(* IEC 61131-3 sources: axsharp/src/AXSharp.connectors/tests/ax-test-project/src, 12 files *)

(* ---- enum.st ---- *)
TYPE
    Colors : (RED, GREEN, BLUE);
END_TYPE

(* ---- complexArrayItem.st ---- *)
{S7.extern=ReadWrite}
CLASS complexArrayItem
    VAR PUBLIC
        itemBOOL	        :       BOOL	      ;
        itemSTRING	        :   STRING	      ;
        itemINT	    :       INT	      ;

    END_VAR
END_CLASS

(* ---- complexArrayItemNested.st ---- *)
{S7.extern=ReadWrite}
CLASS complexArrayItemNested
    VAR PUBLIC
        nesteditemBOOL	        :       BOOL	      ;
        nesteditemSTRING	        :   STRING	      ;
        nesteditemINT	    :       INT	      ;
        nestedComplex: complexArrayItem;
    END_VAR
END_CLASS

(* ---- full_of_primitives.st ---- *)
{S7.extern=ReadWrite}
CLASS full_of_primitives
    VAR PUBLIC
        myBOOL	        :       BOOL	      ;
        myBYTE	        :       BYTE	      ;
        myWORD	        :       WORD	      ;
        myDWORD	        :       DWORD	      ;
        myLWORD	        :       LWORD	      ;
        mySINT	        :       SINT	      ;
        myINT	          :       INT	        ;
        myDINT	        :       DINT	      ;
        myLINT	        :       LINT	      ;
        myUSINT	        :       USINT	      ;
        myUINT	        :       UINT	      ;
        myUDINT	        :       UDINT	      ;
        myULINT	        :       ULINT	      ;
        myREAL	        :       REAL	      ;
        myLREAL	        :       LREAL	      ;
        myTIME	        :       TIME	      ;
        myLTIME	        :       LTIME	      ;
        myDATE	        :       DATE	      ;
        myLDATE	        :       LDATE	      ;
        myTIME_OF_DAY	:       TIME_OF_DAY	  ;
        myLTIME_OF_DAY	:       LTIME_OF_DAY  ;
        myDATE_AND_TIME  :      DATE_AND_TIME ;
        myLDATE_AND_TIME :      LDATE_AND_TIME;
        myCHAR	        :       CHAR	      ;
        myWCHAR	        :       WCHAR	      ;
         mySTRING	        :   STRING	      ;
         myWSTRING	    :       WSTRING	      ;
    END_VAR
END_CLASS

(* ---- full_of_primitives_match.st ---- *)
{S7.extern=ReadWrite}
CLASS full_of_primitives_match
    VAR PUBLIC

        myBOOL	            : BOOL;
        myBYTE	            : BOOL;
        myWORD	            : BOOL;
        myDWORD	        : BOOL;
        myLWORD	        : BOOL;
        mySINT	            : BOOL;
        myINT	            : BOOL;
        myDINT	            : BOOL;
        myLINT	            : BOOL;
        myUSINT	        : BOOL;
        myUINT	            : BOOL;
        myUDINT	        : BOOL;
        myULINT	        : BOOL;
        myREAL	            : BOOL;
        myLREAL	        : BOOL;
        myTIME	            : BOOL;
        myLTIME	        : BOOL;
        myDATE	            : BOOL;
        myLDATE	        : BOOL;
        myTIME_OF_DAY	    : BOOL;
        myLTIME_OF_DAY	    : BOOL;
        myDATE_AND_TIME    : BOOL;
        myLDATE_AND_TIME   : BOOL;
        myCHAR	            : BOOL;
        myWCHAR	        : BOOL;
        mySTRING	        : BOOL;
        myWSTRING	        : BOOL;
    END_VAR
END_CLASS

(* ---- hierarchy.st ---- *)
{S7.extern=ReadWrite}
CLASS hierarchy
    VAR PUBLIC
        item  :      hierarchy_2;
    END_VAR
END_CLASS

(* ---- hierarchy_0.st ---- *)
{S7.extern=ReadWrite}
CLASS hierarchy_0
    VAR PUBLIC
        item_member_property_1   :     full_of_primitives;
        item_member_property_2   :     full_of_primitives;
        item_member_property_3   :     full_of_primitives;
        item_member_property_4   :     full_of_primitives;
        item_member_property_5   :     full_of_primitives;
        item_member_property_6   :     full_of_primitives;
        item_member_property_7   :     full_of_primitives;
        item_member_property_8   :     full_of_primitives;
        item_member_property_9   :     full_of_primitives;
        item_member_property_10  :     full_of_primitives;
        item_member_property_12  :     full_of_primitives;
        item_member_property_13  :     full_of_primitives;
        item_member_property_14  :     full_of_primitives;
        item_member_property_15  :     full_of_primitives;
        item_member_property_16  :     full_of_primitives;
        item_member_property_17  :     full_of_primitives;
        item_member_property_18  :     full_of_primitives;
        item_member_property_19  :     full_of_primitives;
    END_VAR
END_CLASS

(* ---- hierarchy_2.st ---- *)
{S7.extern=ReadWrite}
CLASS hierarchy_2
    VAR PUBLIC
        item_member_property_1   :     hierarchy_0;
        item_member_property_2   :     hierarchy_0;
        item_member_property_3   :     hierarchy_0;
        item_member_property_4   :     hierarchy_0;
        item_member_property_5   :     hierarchy_0;
        item_member_property_6   :     hierarchy_0;
        item_member_property_7   :     hierarchy_0;
        item_member_property_8   :     hierarchy_0;
        item_member_property_9   :     hierarchy_0;
        item_member_property_10  :     hierarchy_0;
        item_member_property_12  :     hierarchy_0;
        item_member_property_13  :     hierarchy_0;
        item_member_property_14  :     hierarchy_0;
        item_member_property_15  :     hierarchy_0;
        item_member_property_16  :     hierarchy_0;
        item_member_property_17  :     hierarchy_0;
        item_member_property_18  :     hierarchy_0;
        item_member_property_19  :     hierarchy_0;
    END_VAR
END_CLASS

(* ---- hierarchy_4.st ---- *)
{S7.extern=ReadWrite}
CLASS hierarchy_4
    VAR PUBLIC
        item_member_property_1   :     hierarchy_2;
        item_member_property_2   :     hierarchy_2;
        item_member_property_3   :     hierarchy_2;
        item_member_property_4   :     hierarchy_2;
        item_member_property_5   :     hierarchy_2;
        item_member_property_6   :     hierarchy_2;
        item_member_property_7   :     hierarchy_2;
        item_member_property_8   :     hierarchy_2;
        item_member_property_9   :     hierarchy_2;
        item_member_property_10  :     hierarchy_2;
        item_member_property_12  :     hierarchy_2;
        item_member_property_13  :     hierarchy_2;
        item_member_property_14  :     hierarchy_2;
        item_member_property_15  :     hierarchy_2;
        item_member_property_16  :     hierarchy_2;
        item_member_property_17  :     hierarchy_2;
        item_member_property_18  :     hierarchy_2;
        item_member_property_19  :     hierarchy_2;
    END_VAR
END_CLASS

(* ---- hierarchy_6.st ---- *)
{S7.extern=ReadWrite}
CLASS hierarchy_6
    VAR PUBLIC
        item_member_property_1  :      hierarchy_4;
        item_member_property_2  :      hierarchy_4;
        item_member_property_3  :      hierarchy_4;
        item_member_property_4  :      hierarchy_4;
        item_member_property_5  :      hierarchy_4;
        item_member_property_6  :      hierarchy_4;
        item_member_property_7   :     hierarchy_4;
        item_member_property_8  :      hierarchy_4;
        item_member_property_9  :      hierarchy_4;
        item_member_property_10  :     hierarchy_4;
        item_member_property_12  :     hierarchy_4;
        item_member_property_13  :     hierarchy_4;
        item_member_property_14  :     hierarchy_4;
        item_member_property_15  :     hierarchy_4;
        item_member_property_16  :     hierarchy_4;
        item_member_property_17  :     hierarchy_4;
        item_member_property_18  :     hierarchy_4;
        item_member_property_19  :     hierarchy_4;
    END_VAR
END_CLASS

(* ---- configuration.st ---- *)
CONFIGURATION MyConfiguration
    TASK Main(Interval := T#1ms, Priority := 1);
    PROGRAM P1 WITH Main: MyProgram;

    VAR_GLOBAL

        //myArrayComplexNested: ARRAY[0..10] OF complexArrayItemNested;

        //myArrayString: ARRAY[0..10] OF STRING;

        // myArrayComplex: ARRAY[0..10] OF complexArrayItem;
        {S7.extern=ReadWrite}
        mins : full_of_primitives;
        {S7.extern=ReadWrite}
        maxs : full_of_primitives;

        {S7.extern=ReadWrite}
        minsmatch : full_of_primitives_match;
        {S7.extern=ReadWrite}
        maxsmatch : full_of_primitives_match;
        {S7.extern=ReadWrite}
        myBOOL	        :       BOOL	 := TRUE     ;
        {S7.extern=ReadWrite}
        myBYTE	        :       BYTE	      ;
        {S7.extern=ReadWrite}
        myWORD	        :       WORD	      ;
        {S7.extern=ReadWrite}
        myDWORD	        :       DWORD	      ;
        {S7.extern=ReadWrite}
        myLWORD	        :       LWORD	      ;
        {S7.extern=ReadWrite}
        mySINT	        :       SINT	      ;
        {S7.extern=ReadWrite}
        myINT	        :       INT	          ;
        {S7.extern=ReadWrite}
        myDINT	        :       DINT	      ;
        {S7.extern=ReadWrite}
        myLINT	        :       LINT	      ;
        {S7.extern=ReadWrite}
        myUSINT	        :       USINT	      ;
        {S7.extern=ReadWrite}
        myUINT	        :       UINT	      ;
        {S7.extern=ReadWrite}
        myUDINT	        :       UDINT	      ;
        {S7.extern=ReadWrite}
        myULINT	        :       ULINT	      ;
        {S7.extern=ReadWrite}
        myREAL	        :       REAL	      ;
        {S7.extern=ReadWrite}
        myLREAL	        :       LREAL	      ;
        {S7.extern=ReadWrite}
        myTIME	        :       TIME	      ;
        {S7.extern=ReadWrite}
        myLTIME	        :       LTIME	      ;
        {S7.extern=ReadWrite}
        myDATE	        :       DATE	      ;
        {S7.extern=ReadWrite}
        myLDATE	        :       LDATE	      ;
        {S7.extern=ReadWrite}
        myTIME_OF_DAY	:       TIME_OF_DAY	  ;
        {S7.extern=ReadWrite}
        myLTIME_OF_DAY	:       LTIME_OF_DAY  ;
        {S7.extern=ReadWrite}
        myDATE_AND_TIME  :      DATE_AND_TIME ;
        {S7.extern=ReadWrite}
        myLDATE_AND_TIME :      LDATE_AND_TIME;
        {S7.extern=ReadWrite}
        myCHAR	        :       CHAR	      ;
        {S7.extern=ReadWrite}
        myWCHAR	        :       WCHAR	      ;
        {S7.extern=ReadWrite}
        mySTRING	        :   STRING	      ;
        {S7.extern=ReadWrite}
        myWSTRING	    :       WSTRING	      ;
        {S7.extern=ReadWrite}
        mySTRING_10	    :       STRING[10]	  ;
        {S7.extern=ReadWrite}
        myWSTRING_10	:       WSTRING[10]	  ;

        {S7.extern=ReadWrite}
        myColors : Colors;

        {S7.extern=ReadWrite}
        Hierarchy : hierarchy;
        // Issues

        //GH_PKTu_ix_56_Base: GH.PKTu.ix_56.Base;

        // GH_PKTu_ix_56_FirstInheritance : GH.PKTu.ix_56.FirstInheritance;
        {S7.extern=ReadWrite}
        GH_PKTu_ix_56_SecondInheritance : GH.PKTu.ix_56.SecondInheritance;

        {S7.extern=ReadWrite}
        myDATE_leap_febr	        :       DATE	      ;
        {S7.extern=ReadWrite}
        myLDATE_leap_febr	        :       LDATE	      ;
        {S7.extern=ReadWrite}
        myDATE_AND_TIME_leap_febr   :      DATE_AND_TIME ;
        {S7.extern=ReadWrite}
        myLDATE_AND_TIME_leap_febr  :      LDATE_AND_TIME;

        {S7.extern=ReadWrite}
        myDATE_leap_late	        :       DATE	      ;
        {S7.extern=ReadWrite}
        myLDATE_leap_late	        :       LDATE	      ;
        {S7.extern=ReadWrite}
        myDATE_AND_TIME_leap_late   :      DATE_AND_TIME ;
        {S7.extern=ReadWrite}
        myLDATE_AND_TIME_leap_late  :      LDATE_AND_TIME;
    END_VAR
END_CONFIGURATION

CONFIGURATION MyConfiguration2
    VAR_GLOBAL
        {S7.extern=ReadWrite}
        mins1 : full_of_primitives;
    END_VAR
END_CONFIGURATION

(* ---- program.st ---- *)
PROGRAM MyProgram
    VAR_EXTERNAL

        //myArrayComplexNested: ARRAY[0..10] OF complexArrayItemNested;

        myBOOL	        :       BOOL	      ;
        myBYTE	        :       BYTE	      ;
        myWORD	        :       WORD	      ;
        myDWORD	        :       DWORD	      ;
        myLWORD	        :       LWORD	      ;
        mySINT	        :       SINT	      ;
        myINT	        :       INT	          ;
        myDINT	        :       DINT	      ;
        myLINT	        :       LINT	      ;
        myUSINT	        :       USINT	      ;
        myUINT	        :       UINT	      ;
        myUDINT	        :       UDINT	      ;
        myULINT	        :       ULINT	      ;
        myREAL	        :       REAL	      ;
        myLREAL	        :       LREAL	      ;
        myTIME	        :       TIME	      ;
        myLTIME	        :       LTIME	      ;
        myDATE	        :       DATE	      ;
        myLDATE	        :       LDATE	      ;
        myTIME_OF_DAY	:       TIME_OF_DAY	  ;
        myLTIME_OF_DAY	:       LTIME_OF_DAY  ;
        myDATE_AND_TIME  :      DATE_AND_TIME ;
        myLDATE_AND_TIME :      LDATE_AND_TIME;
        myCHAR	        :       CHAR	      ;
        myWCHAR	        :       WCHAR	      ;
        mySTRING	        :   STRING	      ;
        myWSTRING	    :       WSTRING	      ;

        mins : full_of_primitives;
        maxs : full_of_primitives;

        minsmatch : full_of_primitives_match;
        maxsmatch : full_of_primitives_match;

        myColors : Colors;

        Hierarchy : hierarchy;

        myDATE_leap_febr	        :       DATE	      ;
        myLDATE_leap_febr	        :       LDATE	      ;
        myDATE_AND_TIME_leap_febr   :      DATE_AND_TIME ;
        myLDATE_AND_TIME_leap_febr  :      LDATE_AND_TIME;

        myDATE_leap_late	        :       DATE	      ;
        myLDATE_leap_late	        :       LDATE	      ;
        myDATE_AND_TIME_leap_late   :      DATE_AND_TIME ;
        myLDATE_AND_TIME_leap_late  :      LDATE_AND_TIME;
        //myArrayString: ARRAY[0..10] OF STRING ;
        //myArrayComplex: ARRAY[0..10] OF complexArrayItem;

    END_VAR

    VAR
        _item : complexArrayItem;
    END_VAR

    VAR_TEMP

    END_VAR

    //myArrayComplex[1] :=  _item;
    //myArrayString[1] := 'ahoj2';

    //myDATE := DATE#2025-02-27;
    //myColors := Colors#GREEN;
    //mins.myBOOL	            :=  false    ;
    mins.myBYTE	            :=  BYTE#2#0    ;
    mins.myWORD	            :=  WORD#0    ;
    mins.myDWORD	        :=  DWORD#16#0    ;
    mins.myLWORD	        :=  LWORD#0    ;
    mins.mySINT	            :=  SINT#-128    ;
    mins.myINT	            :=  INT#-32768      ;
    mins.myDINT	            :=  DINT#-2147483648;
    mins.myLINT	            :=  LINT#-9223372036854775808    ;
    mins.myUSINT	        :=  USINT#0    ;
    mins.myUINT	            :=  UINT#0    ;
    mins.myUDINT	        :=  UDINT#0     ;
    mins.myULINT	        :=  ULINT#0    ;
    mins.myREAL	            :=  REAL#-3.402823e+38    ;
    mins.myLREAL	        :=  LREAL#-1.79769313486231e+308;
    mins.myTIME	            :=  TIME#-106751d23h47m16s854ms;
    mins.myLTIME	        :=  LTIME#-106751d23h47m16s854ms;
    mins.myDATE	            :=  DATE#1970-01-01    ;
    mins.myLDATE	        :=  LDATE#1970-01-01    ;
    mins.myTIME_OF_DAY	    :=  TOD#0:0:0.0   ;
    mins.myLTIME_OF_DAY	    :=  LTOD#0:0:0.0    ;
    mins.myDATE_AND_TIME    :=  DT#1970-01-01-0:0:0.0   ;
    mins.myLDATE_AND_TIME   :=  LDT#1970-01-01-0:0:0.0   ;
    mins.myCHAR	            :=  CHAR#' '    ;
    mins.myWCHAR	        :=  WCHAR#" "    ;
    mins.mySTRING	        :=  STRING#'';
    mins.myWSTRING	        :=  WSTRING#""    ;

    maxs.myBOOL	            :=  TRUE    ;
    maxs.myBYTE	            :=  BYTE#255    ;
    maxs.myWORD	            :=  WORD#065535    ;
    maxs.myDWORD	        :=  DWORD#4294967295    ;
    maxs.myLWORD	        :=  LWORD#18446744073709551615    ;
    maxs.mySINT	            :=  SINT#127    ;
    maxs.myINT	            :=  INT#32767      ;
    maxs.myDINT	            :=  DINT#2147483647;
    maxs.myLINT	            :=  LINT#9223372036854775807    ;
    maxs.myUSINT	        :=  USINT#255    ;
    maxs.myUINT	            :=  UINT#65535    ;
    maxs.myUDINT	        :=  UDINT#4294967295     ;
    maxs.myULINT	        :=  ULINT#18446744073709551615    ;
    maxs.myREAL	            :=  REAL#+3.402823e+38    ;
    maxs.myLREAL	        :=  LREAL#1.79769313486231e+308;
    maxs.myTIME	            :=  TIME#106751d23h47m16s854ms;
    maxs.myLTIME	        :=  LTIME#106751d23h47m16s854ms;
    maxs.myLTIME	        :=  LTIME#106751d23h47m16s854ms;
    // maxs.myLTIME	        :=  LTIME#1067d12h28m40s368ms547us758ns;
    maxs.myDATE	            :=  DATE#2262-04-11    ;
    maxs.myLDATE	        :=  LDATE#2262-04-11    ;
    maxs.myTIME_OF_DAY	    :=  TOD#23:59:59.999000000   ;
    maxs.myLTIME_OF_DAY	    :=  LTOD#23:59:59.999000000    ;
    maxs.myDATE_AND_TIME    :=  DT#2262-04-11-23:47:16.854   ;
    maxs.myLDATE_AND_TIME   :=  LDT#2262-04-11-23:47:16.854   ;
    maxs.myCHAR	            :=  CHAR#'$7F';
    maxs.myWCHAR	        :=  WCHAR#"$D7FE";
    maxs.mySTRING	        :=  STRING#'ABCDEFGHIJKLMNOPRSTUABCDEFGHIJKLMNOPRSTUABCDEFGHIJKLMNOPRSTUABCDEFGHIJKLMNOPRSTUABCDEFGHIJKLMNOPRSTUABCDEFGHIJKLMNOPRSTUABCDEFGHIJKLMNOPRSTUABCDEFGHIJKLMNOPRSTUABCDEFGHIJKLMNOPRSTUABCDEFGHIJKLMNOPRSTUABCDEFGHIJKLMNOPRSTUABCDEFGHIJKLMNOPRSTUABCDEFGHIJKLMN';
    maxs.myWSTRING	        :=  WSTRING#"ABCDEFGHIJKLMNOPRSTUABCDEFGHIJKLMNOPRSTUABCDEFGHIJKLMNOPRSTUABCDEFGHIJKLMNOPRSTUABCDEFGHIJKLMNOPRSTUABCDEFGHIJKLMNOPRSTUABCDEFGHIJKLMNOPRSTUABCDEFGHIJKLMNOPRSTUABCDEFGHIJKLMNOPRSTUABCDEFGHIJKLMNOPRSTUABCDEFGHIJKLMNOPRSTUABCDEFGHIJKLMNOPRSTUABCDEFGHIJKLMN";

    minsmatch.myBOOL	        := mins.myBOOL	         =  myBOOL	        ;
    minsmatch.myBYTE	        := mins.myBYTE	         =  myBYTE	        ;
    minsmatch.myWORD	        := mins.myWORD	         =  myWORD	        ;
    minsmatch.myDWORD	        := mins.myDWORD	         =  myDWORD	        ;
    minsmatch.myLWORD	        := mins.myLWORD	         =  myLWORD	        ;
    minsmatch.mySINT	        := mins.mySINT	         =  mySINT	        ;
    minsmatch.myINT	            := mins.myINT	         =  myINT	        ;
    minsmatch.myDINT	        := mins.myDINT	         =  myDINT	        ;
    minsmatch.myLINT	        := mins.myLINT	         =  myLINT	        ;
    minsmatch.myUSINT	        := mins.myUSINT	         =  myUSINT	        ;
    minsmatch.myUINT	        := mins.myUINT	         =  myUINT	        ;
    minsmatch.myUDINT	        := mins.myUDINT	         =  myUDINT	        ;
    minsmatch.myULINT	        := mins.myULINT	         =  myULINT	        ;
    minsmatch.myREAL	        := mins.myREAL	         =  myREAL	        ;
    minsmatch.myLREAL	        := mins.myLREAL	         =  myLREAL	        ;
    minsmatch.myTIME	        := mins.myTIME	         =  myTIME	        ;
    minsmatch.myLTIME	        := mins.myLTIME	         =  myLTIME	        ;
    minsmatch.myDATE	        := mins.myDATE	         =  myDATE	        ;
    minsmatch.myLDATE	        := mins.myLDATE	         =  myLDATE	        ;
    minsmatch.myTIME_OF_DAY	    := mins.myTIME_OF_DAY	 =  myTIME_OF_DAY	;
    minsmatch.myLTIME_OF_DAY	:= mins.myLTIME_OF_DAY	 =  myLTIME_OF_DAY	;
    minsmatch.myDATE_AND_TIME   := mins.myDATE_AND_TIME  =  myDATE_AND_TIME ;
    minsmatch.myLDATE_AND_TIME  := mins.myLDATE_AND_TIME =  myLDATE_AND_TIME;
    minsmatch.myCHAR	        := mins.myCHAR	         =  myCHAR	        ;
    minsmatch.myWCHAR	        := mins.myWCHAR	         =  myWCHAR	        ;
    minsmatch.mySTRING	        := mins.mySTRING	     =  mySTRING	    ;
    minsmatch.myWSTRING	        := mins.myWSTRING	     =  myWSTRING	    ;

    maxsmatch.myBOOL	        := maxs.myBOOL	         =  myBOOL	        ;
    maxsmatch.myBYTE	        := maxs.myBYTE	         =  myBYTE	        ;
    maxsmatch.myWORD	        := maxs.myWORD	         =  myWORD	        ;
    maxsmatch.myDWORD	        := maxs.myDWORD	         =  myDWORD	        ;
    maxsmatch.myLWORD	        := maxs.myLWORD	         =  myLWORD	        ;
    maxsmatch.mySINT	        := maxs.mySINT	         =  mySINT	        ;
    maxsmatch.myINT	            := maxs.myINT	         =  myINT	        ;
    maxsmatch.myDINT	        := maxs.myDINT	         =  myDINT	        ;
    maxsmatch.myLINT	        := maxs.myLINT	         =  myLINT	        ;
    maxsmatch.myUSINT	        := maxs.myUSINT	         =  myUSINT	        ;
    maxsmatch.myUINT	        := maxs.myUINT	         =  myUINT	        ;
    maxsmatch.myUDINT	        := maxs.myUDINT	         =  myUDINT	        ;
    maxsmatch.myULINT	        := maxs.myULINT	         =  myULINT	        ;
    maxsmatch.myREAL	        := maxs.myREAL	         =  myREAL	        ;
    maxsmatch.myLREAL	        := maxs.myLREAL	         =  myLREAL	        ;
    maxsmatch.myTIME	        := maxs.myTIME	         =  myTIME	        ;
    maxsmatch.myLTIME	        := maxs.myLTIME	         =  myLTIME	        ;
    maxsmatch.myDATE	        := maxs.myDATE	         =  myDATE	        ;
    maxsmatch.myLDATE	        := maxs.myLDATE	         =  myLDATE	        ;
    maxsmatch.myTIME_OF_DAY	    := maxs.myTIME_OF_DAY	 =  myTIME_OF_DAY	;
    maxsmatch.myLTIME_OF_DAY	:= maxs.myLTIME_OF_DAY	 =  myLTIME_OF_DAY	;
    maxsmatch.myDATE_AND_TIME   := maxs.myDATE_AND_TIME  =  myDATE_AND_TIME ;
    maxsmatch.myLDATE_AND_TIME  := maxs.myLDATE_AND_TIME =  myLDATE_AND_TIME;
    maxsmatch.myCHAR	        := maxs.myCHAR	         =  myCHAR	        ;
    maxsmatch.myWCHAR	        := maxs.myWCHAR	         =  myWCHAR	        ;
    maxsmatch.mySTRING	        := maxs.mySTRING	     =  mySTRING	    ;
    maxsmatch.myWSTRING	        := maxs.myWSTRING	     =  myWSTRING	    ;

    myDATE_leap_febr	        :=  DATE#2024-02-29;
    myLDATE_leap_febr	        :=  LDATE#2024-02-29;
    myDATE_AND_TIME_leap_febr   :=  DATE_AND_TIME#2024-02-29-0:0:0.0;
    myLDATE_AND_TIME_leap_febr  :=  LDATE_AND_TIME#2024-02-29-0:0:0.0;

    myDATE_leap_late	        :=   DATE#2024-03-05;
    myLDATE_leap_late	        :=   LDATE#2024-03-05;
    myDATE_AND_TIME_leap_late   :=   DATE_AND_TIME#2024-03-05-0:0:0.0;
    myLDATE_AND_TIME_leap_late  :=   LDATE_AND_TIME#2024-03-05-0:0:0.0;
END_PROGRAM
